(* IEC 61131-3 sources: plc-process-lib/tests/POUs/Suites/FB_DeviceBase_Test, 53 files *)

(* ---- AckAllAcksEveryAlarm.method.decl.st ---- *)
// AckAll() квитирует все тревоги устройства: три активных слота → ActiveAck, wAlmUnack = 0, бит
// DEV_STS_ALARM_UNACK снят, результат Accepted; когда квитировать нечего, AckAll() — FALSE.
// Бит stCmd.xAck делает то же и сбрасывается.
METHOD PRIVATE AckAllAcksEveryAlarm
VAR
    fbTime   : FB_FakeTime;        // подменное время
    fbDev    : FB_TestDevice;      // устройство под тестом
    stCmd    : ST_TestDeviceCmd;   // команды
    stRetain : ST_DeviceRetain;    // энергонезависимые данные
    stCfg    : ST_TestDeviceCfg;   // конфигурация по умолчанию
    itfAlm   : I_Alarm;            // слот через интерфейс
    xRet     : BOOL;               // ответ AckAll
END_VAR

(* ---- AckMaskAcksOnlySelectedSlot.method.decl.st ---- *)
// Маска wAckReq квитирует только выбранный слот (бит 1), маска обнуляется, результат Accepted.
METHOD PRIVATE AckMaskAcksOnlySelectedSlot
VAR
    fbTime   : FB_FakeTime;        // подменное время
    fbDev    : FB_TestDevice;      // устройство под тестом
    stCmd    : ST_TestDeviceCmd;   // команды
    stRetain : ST_DeviceRetain;    // энергонезависимые данные
    stCfg    : ST_TestDeviceCfg;   // конфигурация по умолчанию
    itfAlm   : I_Alarm;            // слот через интерфейс
END_VAR

(* ---- AlarmIdsBaseFromCfgPlusSlot.method.decl.st ---- *)
// Номер тревоги слота = stCfg.udiAlarmIdBase + слот: база 120, слот 5 — 125; номер и значение
// процесса приходят в событии.
METHOD PRIVATE AlarmIdsBaseFromCfgPlusSlot
VAR
    fbTime   : FB_FakeTime;        // подменное время
    fbDev    : FB_TestDevice;      // устройство под тестом
    stCmd    : ST_TestDeviceCmd;   // команды
    stRetain : ST_DeviceRetain;    // энергонезависимые данные
    stCfg    : ST_TestDeviceCfg;   // udiAlarmIdBase = 120
    fbSink   : FB_TestSink;        // приёмник событий
    stEv     : ST_AlarmEvent;      // последнее событие
    itfAlm   : I_Alarm;            // слот через интерфейс
END_VAR

(* ---- AlarmPriorityInvalidCfgErrBit.method.decl.st ---- *)
// Приоритет тревоги вне перечисления (9) не проходит CheckAlarmCfg: бит wCfgErr устройства и
// CheckFunction; исправленный приоритет снимает бит.
METHOD PRIVATE AlarmPriorityInvalidCfgErrBit
VAR
    fbTime   : FB_FakeTime;        // подменное время
    fbDev    : FB_TestDevice;      // устройство под тестом
    stCmd    : ST_TestDeviceCmd;   // команды
    stRetain : ST_DeviceRetain;    // энергонезависимые данные
    stCfg    : ST_TestDeviceCfg;   // слот 3: приоритет 9
    uBad     : U_TestEnumInt;      // число вне перечисления
END_VAR

(* ---- AlarmsInOosAllSlotsOutOfService.method.decl.st ---- *)
// OutOfService устройства — OutOfService у всех используемых слотов (3); в wAlmShelved и wAlmSuppressed их нет
// (ALM-2: вывод из работы виден по eMode), неквитированных нет; после выхода активная тревога снова ActiveUnack.
METHOD PRIVATE AlarmsInOosAllSlotsOutOfService
VAR
    fbTime   : FB_FakeTime;        // подменное время
    fbDev    : FB_TestDevice;      // устройство под тестом
    stCmd    : ST_TestDeviceCmd;   // команды
    stRetain : ST_DeviceRetain;    // энергонезависимые данные
    stCfg    : ST_TestDeviceCfg;   // конфигурация по умолчанию
    itfAlm   : I_Alarm;            // слот через интерфейс
END_VAR

(* ---- AlarmSlotArraysMatchDevAlarmsMax.method.decl.st ---- *)
// Длина массивов слотов базы (afbAlarm, axAlmCond, axAlmSuppress, arAlmValue) равна
// GVL_Const.DEV_ALARMS_MAX: циклы базы идут по константе, тест ловит расхождение, если границу
// запишут числом. Тест читает внутренние переменные базы намеренно — это проверка раскладки.
METHOD PRIVATE AlarmSlotArraysMatchDevAlarmsMax
VAR
    fbDev : FB_TestDevice;   // устройство (вызов не нужен)
    fbAlm : FB_Alarm;        // размер одного слота
END_VAR

(* ---- AlarmSummaryWordsAndPrioUnack.method.decl.st ---- *)
// Сводка тревог: слоты Low, High, Medium активны — ePrioUnack = High; квитирован High — Medium;
// слот Medium вернулся без квитирования — wAlmActive = 2#011, wAlmUnack = 2#101; подавление слота 0
// — бит в wAlmSuppressed (не в wAlmShelved, ALM-2) и снят из wAlmUnack.
METHOD PRIVATE AlarmSummaryWordsAndPrioUnack
VAR
    fbTime   : FB_FakeTime;        // подменное время
    fbDev    : FB_TestDevice;      // устройство под тестом
    stCmd    : ST_TestDeviceCmd;   // команды
    stRetain : ST_DeviceRetain;    // энергонезависимые данные
    stCfg    : ST_TestDeviceCfg;   // приоритеты слотов 0…2
END_VAR

(* ---- AutoToManualBumplessKeepsOutput.method.decl.st ---- *)
// Безударный переход Auto → Manual (хук наследника): работающий механизм продолжает работать.
METHOD PRIVATE AutoToManualBumplessKeepsOutput
VAR
    fbTime   : FB_FakeTime;        // подменное время
    fbDev    : FB_TestDevice;      // устройство под тестом
    stCmd    : ST_TestDeviceCmd;   // команды
    stRetain : ST_DeviceRetain;    // энергонезависимые данные
    stCfg    : ST_TestDeviceCfg;   // конфигурация по умолчанию
END_VAR

(* ---- BeginCycleDtZeroOnFirstCallThenFromTimeSource.method.decl.st ---- *)
// BeginCycle: в первом вызове ltDt = 0; затем — шаг подменного времени (250 мс); при «времени
// назад» — 0 (без переполнения LTIME); дальше снова шаг (100 мс).
METHOD PRIVATE BeginCycleDtZeroOnFirstCallThenFromTimeSource
VAR
    fbTime   : FB_FakeTime;        // подменное время
    fbDev    : FB_TestDevice;      // устройство под тестом
    stCmd    : ST_TestDeviceCmd;   // команды
    stRetain : ST_DeviceRetain;    // энергонезависимые данные
    stCfg    : ST_TestDeviceCfg;   // конфигурация по умолчанию
END_VAR

(* ---- CmdBitsClearedAfterProcessing.method.decl.st ---- *)
// Все импульсные биты и маски stCmd (xSetAuto, xSetManual, xSetOos, xReset, xAck, wAckReq,
// wShelveReq, wUnshelveReq, xStart, xStop) сброшены в том же вызове.
METHOD PRIVATE CmdBitsClearedAfterProcessing
VAR
    fbTime   : FB_FakeTime;        // подменное время
    fbDev    : FB_TestDevice;      // устройство под тестом
    stCmd    : ST_TestDeviceCmd;   // команды
    stRetain : ST_DeviceRetain;    // энергонезависимые данные
    stCfg    : ST_TestDeviceCfg;   // конфигурация по умолчанию
END_VAR

(* ---- CmdResultSeqIncrementsPerCommand.method.decl.st ---- *)
// Каждая обработанная команда пишет eCmdResult и увеличивает uiCmdSeq: в одном вызове режим и пуск
// (в Auto отклонён) — +2, результат последней RejectedMode; Reset и маска shelve без
// принявших слотов — +2, результат RejectedState.
METHOD PRIVATE CmdResultSeqIncrementsPerCommand
VAR
    fbTime   : FB_FakeTime;        // подменное время
    fbDev    : FB_TestDevice;      // устройство под тестом
    stCmd    : ST_TestDeviceCmd;   // команды
    stRetain : ST_DeviceRetain;    // энергонезависимые данные
    stCfg    : ST_TestDeviceCfg;   // слот 0: shelve запрещён
END_VAR

(* ---- ConflictingModeRequestsOosWins.method.decl.st ---- *)
// Одновременные запросы режима (xSetAuto, xSetManual, xSetOos и RequestMode(Auto)) — одна команда:
// побеждает OutOfService; затем xSetAuto вместе с RequestMode(Manual) — побеждает Manual и выводит
// из OutOfService. Импульсы сброшены.
METHOD PRIVATE ConflictingModeRequestsOosWins
VAR
    fbTime   : FB_FakeTime;        // подменное время
    fbDev    : FB_TestDevice;      // устройство под тестом
    stCmd    : ST_TestDeviceCmd;   // команды
    stRetain : ST_DeviceRetain;    // энергонезависимые данные
    stCfg    : ST_TestDeviceCfg;   // конфигурация по умолчанию
    xRet     : BOOL;               // ответ RequestMode
END_VAR

(* ---- DefaultAlarmCfgOfAllTypesPassesCheckAlarmCfg.method.decl.st ---- *)
// Умолчания astAlarm Cfg всех семи устройств и тестового проходят CheckAlarmCfg (инвариант
// генератора для конфигурации тревог); массивы astAlarm из DUT передаются в параметр
// ARRAY[0..GVL_Const.DEV_ALARMS_MAX - 1]. Приоритет 5 и -1 — отказ, 4 (Critical) — норма.
METHOD PRIVATE DefaultAlarmCfgOfAllTypesPassesCheckAlarmCfg
VAR
    fbDev  : FB_TestDevice;         // доступ к CheckAlarmCfg
    stAi   : ST_AnalogInputCfg;     // умолчания AI
    stDi   : ST_DigitalInputCfg;    // умолчания DI
    stMot  : ST_MotorCfg;           // умолчания двигателя
    stVlv  : ST_ValveCfg;           // умолчания арматуры
    stCv   : ST_ControlValveCfg;    // умолчания регулирующего клапана
    stPid  : ST_PidCfg;             // умолчания ПИД
    stTest : ST_TestDeviceCfg;      // умолчания тестового устройства
    stSlot : ST_AlarmCfg;           // копия слота
    uBad   : U_TestEnumInt;         // число вне перечисления
END_VAR

(* ---- DerivedBodyWithoutSuperBaseBodyNotRun.method.decl.st ---- *)
// L1 контракта во время выполнения: у наследника со своим телом без SUPER^ тело базы не
// выполняется само — импульс режима не обработан, FinishCycle не вызван (eDevType = None).
METHOD PRIVATE DerivedBodyWithoutSuperBaseBodyNotRun
VAR
    fbTime   : FB_FakeTime;            // подменное время
    fbNo     : FB_TestDeviceNoSuper;   // наследник без SUPER^
    stCmd    : ST_TestDeviceCmd;       // команды
    stRetain : ST_DeviceRetain;        // энергонезависимые данные
    stCfg    : ST_TestDeviceCfg;       // конфигурация по умолчанию
END_VAR

(* ---- DevTypeSetByHeirReportedInStsCommon.method.decl.st ---- *)
// Тип устройства задаёт наследник в первом вызове, FinishCycle пишет его в stCommon.eDevType;
// до первого вызова — None.
METHOD PRIVATE DevTypeSetByHeirReportedInStsCommon
VAR
    fbTime   : FB_FakeTime;        // подменное время
    fbDev    : FB_TestDevice;      // устройство под тестом
    stCmd    : ST_TestDeviceCmd;   // команды
    stRetain : ST_DeviceRetain;    // энергонезависимые данные
    stCfg    : ST_TestDeviceCfg;   // конфигурация по умолчанию
END_VAR

(* ---- FailureSafeStateResetRules.method.decl.st ---- *)
// Безопасное состояние при отказе: выход снят, Fault, NE 107 Failure, бит wFault, Available =
// FALSE. Reset при действующей причине — RejectedFault; причина ушла — отказ держится до Reset();
// после Reset() выход не включается сам (ручная защёлка снята).
METHOD PRIVATE FailureSafeStateResetRules
VAR
    fbTime   : FB_FakeTime;        // подменное время
    fbDev    : FB_TestDevice;      // устройство под тестом
    stCmd    : ST_TestDeviceCmd;   // команды
    stRetain : ST_DeviceRetain;    // энергонезависимые данные
    stCfg    : ST_TestDeviceCfg;   // конфигурация по умолчанию
    xRet     : BOOL;               // ответ Reset
END_VAR

(* ---- GetAlarmOutOfRangeReturnsNull.method.decl.st ---- *)
// GetAlarm отдаёт слот только в 0..AlarmCount - 1: при трёх слотах — слоты 0…2, номер 3 и 65535 —
// 0; до первого вызова слотов нет.
METHOD PRIVATE GetAlarmOutOfRangeReturnsNull
VAR
    fbTime   : FB_FakeTime;        // подменное время
    fbDev    : FB_TestDevice;      // устройство под тестом
    stCmd    : ST_TestDeviceCmd;   // команды
    stRetain : ST_DeviceRetain;    // энергонезависимые данные
    stCfg    : ST_TestDeviceCfg;   // конфигурация по умолчанию
    itfAlm   : I_Alarm;            // ответ GetAlarm
END_VAR

(* ---- HookViaThisDispatchesToMostDerivedOverride.method.decl.st ---- *)
// Вопрос R2 для двух уровней: у FB_TestDeviceExt хук переопределён ещё раз. THIS^.OnModeChanged из
// метода FB_DeviceBase вызывает реализацию самого производного ФБ; её SUPER^.OnModeChanged
// выполняет часть FB_TestDevice, затем своя часть: след 12 на одну смену режима, 1212 — на две.
METHOD PRIVATE HookViaThisDispatchesToMostDerivedOverride
VAR
    fbTime   : FB_FakeTime;        // подменное время
    fbExt    : FB_TestDeviceExt;   // наследник второго уровня
    stCmd    : ST_TestDeviceCmd;   // команды
    stRetain : ST_DeviceRetain;    // энергонезависимые данные
    stCfg    : ST_TestDeviceCfg;   // конфигурация по умолчанию
END_VAR

(* ---- ImplementsIDeviceInterfaceAccess.method.decl.st ---- *)
// Устройства через I_Device (массив интерфейсов, как у станционной логики): RequestMode, Reset,
// Mode, Status, Fault, Available, AlarmCount, GetAlarm, AckAll работают одинаково для
// FB_TestDevice и его наследника.
METHOD PRIVATE ImplementsIDeviceInterfaceAccess
VAR
    fbTime    : FB_FakeTime;        // подменное время
    fbDev     : FB_TestDevice;      // первое устройство
    fbExt     : FB_TestDeviceExt;   // второе устройство (наследник)
    stCmd     : ST_TestDeviceCmd;   // команды первого
    stRetain  : ST_DeviceRetain;    // retain первого
    stCmd2    : ST_TestDeviceCmd;   // команды второго
    stRetain2 : ST_DeviceRetain;    // retain второго
    stCfg     : ST_TestDeviceCfg;   // общая конфигурация
    aitfDev   : ARRAY[0..1] OF I_Device;   // устройства через интерфейс
    itfDev    : I_Device;           // элемент массива
    itfAlm    : I_Alarm;            // тревога через интерфейс
    uiDev     : UINT;               // номер устройства
    xAllAuto  : BOOL := TRUE;       // все в Auto
    xRet      : BOOL;               // ответы методов
END_VAR

(* ---- ImplementsIDeviceInterfaceAccess.method.impl.st ---- *)
coUnit.TEST('Device_ImplementsIDevice_InterfaceAccess');

aitfDev[0] := fbDev;
aitfDev[1] := fbExt;
FOR uiDev := 0 TO 1 DO
    itfDev := aitfDev[uiDev];
    itfDev.RequestMode(eNewMode := E_DeviceMode.Auto);
END_FOR
fbDev.axCondIn[0] := TRUE;
fbDev(xFaultCause := TRUE, itfTime := fbTime, stCmd := stCmd, stRetain := stRetain, stCfg := stCfg);
fbExt(itfTime := fbTime, stCmd := stCmd2, stRetain := stRetain2, stCfg := stCfg);
FOR uiDev := 0 TO 1 DO
    itfDev := aitfDev[uiDev];
    xAllAuto := xAllAuto AND itfDev.Mode = E_DeviceMode.Auto;
END_FOR
AssertTrue(Condition := xAllAuto, Message := 'RequestMode through the interface');
itfDev := aitfDev[0];
AssertTrue(Condition := itfDev.Fault, Message := 'Fault through the interface');
AssertTrue(Condition := itfDev.Status = E_Ne107Status.Failure, Message := 'Status through the interface');
AssertFalse(Condition := itfDev.Available, Message := 'Available through the interface');
AssertEquals_UINT(Expected := 8, Actual := itfDev.AlarmCount, Message := 'AlarmCount through the interface');
itfAlm := itfDev.GetAlarm(uiIndex := 0);
AssertTrue(Condition := itfAlm.Unacked, Message := 'GetAlarm through the interface');
xRet := itfDev.AckAll();
AssertTrue(Condition := xRet, Message := 'AckAll through the interface');
itfDev.Reset();
fbDev(xFaultCause := FALSE, itfTime := fbTime, stCmd := stCmd, stRetain := stRetain, stCfg := stCfg);
AssertFalse(Condition := itfDev.Fault, Message := 'Reset through the interface');
AssertFalse(Condition := itfAlm.Unacked, Message := 'alarm acknowledged');
itfDev := aitfDev[1];
AssertTrue(Condition := itfDev.Available, Message := 'second device available in Auto');

coUnit.TEST_FINISHED();

(* ---- InputLikeModeMemStartsAutoManualIsCheck.method.decl.st ---- *)
// AI/DI-подобное устройство (без stRetain, режима Local нет): после старта Auto из stModeMem,
// переключатель «Местное» не действует, xSetManual — Manual (подмена) с CheckFunction; stRetain не
// трогается.
METHOD PRIVATE InputLikeModeMemStartsAutoManualIsCheck
VAR
    fbTime   : FB_FakeTime;        // подменное время
    fbIn     : FB_TestDevice;      // устройство под тестом
    stCmd    : ST_TestDeviceCmd;   // команды
    stRetain : ST_DeviceRetain;    // не используется
    stCfg    : ST_TestDeviceCfg;   // конфигурация по умолчанию
END_VAR

(* ---- InvalidCfgAtStartCheckFunctionSafeOutput.method.decl.st ---- *)
// Корректной Cfg ещё не было (rGain = 0): бит wCfgErr, NE 107 CheckFunction, DEV_STS_CFG_ERROR,
// безопасный выход (FALSE и в Auto с запросом), Available = FALSE, пуск — RejectedCfg; режимы
// работают.
METHOD PRIVATE InvalidCfgAtStartCheckFunctionSafeOutput
VAR
    fbTime   : FB_FakeTime;        // подменное время
    fbDev    : FB_TestDevice;      // устройство под тестом
    stCmd    : ST_TestDeviceCmd;   // команды
    stRetain : ST_DeviceRetain;    // энергонезависимые данные
    stCfg    : ST_TestDeviceCfg;   // rGain = 0 — неверно
END_VAR

(* ---- InvalidCfgDuringOperationKeepsLastValidCfg.method.decl.st ---- *)
// Cfg испорчена в работе (rGain = -1): бит wCfgErr и CheckFunction, но логика работает по LKG
// (значение 20 от rGain = 2), механизм не останавливается, Available не меняется; исправленная
// Cfg (rGain = 3) принимается сразу.
METHOD PRIVATE InvalidCfgDuringOperationKeepsLastValidCfg
VAR
    fbTime   : FB_FakeTime;        // подменное время
    fbDev    : FB_TestDevice;      // устройство под тестом
    stCmd    : ST_TestDeviceCmd;   // команды
    stRetain : ST_DeviceRetain;    // энергонезависимые данные
    stCfg    : ST_TestDeviceCfg;   // rGain = 2, затем -1 и 3
END_VAR

(* ---- LocalModeNe107CheckFunction.method.decl.st ---- *)
// Local (переключатель на месте, тип с Local): ПЛК механизмом не управляет — сводный NE 107 CheckFunction («местное
// управление», категория C NE 107, статус PA 0x3C), Available = FALSE; отказ в Local старше — Failure. Возврат в
// дистанционный режим — Good.
METHOD PRIVATE LocalModeNe107CheckFunction
VAR
    fbTime   : FB_FakeTime;        // подменное время
    fbDev    : FB_TestDevice;      // устройство под тестом
    stCmd    : ST_TestDeviceCmd;   // команды
    stRetain : ST_DeviceRetain;    // энергонезависимые данные
    stCfg    : ST_TestDeviceCfg;   // конфигурация
END_VAR

(* ---- LocalOverridesRemoteReturnsToRememberedMode.method.decl.st ---- *)
// Local старше дистанционного режима: в Local выходы сняты, запомненный режим (Auto) сохранён;
// после возврата переключателя устройство продолжает в Auto. Хук — на каждой смене режима.
METHOD PRIVATE LocalOverridesRemoteReturnsToRememberedMode
VAR
    fbTime   : FB_FakeTime;        // подменное время
    fbDev    : FB_TestDevice;      // устройство под тестом
    stCmd    : ST_TestDeviceCmd;   // команды
    stRetain : ST_DeviceRetain;    // энергонезависимые данные
    stCfg    : ST_TestDeviceCfg;   // конфигурация по умолчанию
END_VAR

(* ---- MethodRequestsProcessedOnce.method.decl.st ---- *)
// Запросы методов Reset(), AckAll() и RequestMode() выполняет один ближайший вызов тела, затем они
// снимаются (FinishCycle): uiCmdSeq растёт на 1 за запрос, а не в каждом цикле; тревога, появившаяся
// после выполненного запроса, остаётся неквитированной; режим, сменённый командой после
// RequestMode(), повторный запрос не возвращает. Иначе Reset() станции квитировал бы все будущие
// тревоги и бесконечно повторял бы сброс
METHOD PRIVATE MethodRequestsProcessedOnce
VAR
    fbTime   : FB_FakeTime;        // подменное время
    fbDev    : FB_TestDevice;      // устройство под тестом
    stCmd    : ST_TestDeviceCmd;   // команды
    stRetain : ST_DeviceRetain;    // энергонезависимые данные
    stCfg    : ST_TestDeviceCfg;   // конфигурация по умолчанию
    iStep    : INT;                // шаг цикла
END_VAR

(* ---- MethodRequestsProcessedOnce.method.impl.st ---- *)
coUnit.TEST('Device_MethodRequests_ProcessedOnce');

fbDev(itfTime := fbTime, stCmd := stCmd, stRetain := stRetain, stCfg := stCfg);
fbDev.Reset();
FOR iStep := 1 TO 3 DO
    fbTime.Advance(tStep := T#100MS);
    fbDev(itfTime := fbTime, stCmd := stCmd, stRetain := stRetain, stCfg := stCfg);
END_FOR
AssertEquals_UINT(Expected := 1, Actual := fbDev.stSts.stCommon.uiCmdSeq, Message := 'Reset() executed once');
fbDev.axCondIn[0] := TRUE;
fbDev(itfTime := fbTime, stCmd := stCmd, stRetain := stRetain, stCfg := stCfg);
fbDev(itfTime := fbTime, stCmd := stCmd, stRetain := stRetain, stCfg := stCfg);
AssertEquals_WORD(Expected := 16#0001, Actual := fbDev.stSts.stCommon.wAlmUnack,
                  Message := 'alarm after Reset() stays unacknowledged');
AssertEquals_UINT(Expected := 1, Actual := fbDev.stSts.stCommon.uiCmdSeq, Message := 'no repeated reset');

fbDev.AckAll();
fbDev(itfTime := fbTime, stCmd := stCmd, stRetain := stRetain, stCfg := stCfg);
AssertEquals_WORD(Expected := 0, Actual := fbDev.stSts.stCommon.wAlmUnack, Message := 'AckAll() acknowledged');
fbDev.axCondIn[1] := TRUE;
fbDev(itfTime := fbTime, stCmd := stCmd, stRetain := stRetain, stCfg := stCfg);
fbDev(itfTime := fbTime, stCmd := stCmd, stRetain := stRetain, stCfg := stCfg);
AssertEquals_WORD(Expected := 16#0002, Actual := fbDev.stSts.stCommon.wAlmUnack,
                  Message := 'alarm after AckAll() stays unacknowledged');
AssertEquals_UINT(Expected := 2, Actual := fbDev.stSts.stCommon.uiCmdSeq, Message := 'AckAll() executed once');

fbDev.RequestMode(eNewMode := E_DeviceMode.Auto);
fbDev(itfTime := fbTime, stCmd := stCmd, stRetain := stRetain, stCfg := stCfg);
AssertTrue(Condition := fbDev.Mode = E_DeviceMode.Auto, Message := 'RequestMode(Auto) executed');
stCmd.stCommon.xSetManual := TRUE;
fbDev(itfTime := fbTime, stCmd := stCmd, stRetain := stRetain, stCfg := stCfg);
fbDev(itfTime := fbTime, stCmd := stCmd, stRetain := stRetain, stCfg := stCfg);
AssertTrue(Condition := fbDev.Mode = E_DeviceMode.Manual, Message := 'old RequestMode(Auto) does not come back');
AssertEquals_UINT(Expected := 4, Actual := fbDev.stSts.stCommon.uiCmdSeq, Message := 'four commands in total');

coUnit.TEST_FINISHED();

(* ---- ModeRequestInLocalChangesRememberedMode.method.decl.st ---- *)
// В Local команда xSetAuto принимается и меняет только запомненный режим; после возврата
// переключателя устройство работает в Auto.
METHOD PRIVATE ModeRequestInLocalChangesRememberedMode
VAR
    fbTime   : FB_FakeTime;        // подменное время
    fbDev    : FB_TestDevice;      // устройство под тестом
    stCmd    : ST_TestDeviceCmd;   // команды
    stRetain : ST_DeviceRetain;    // энергонезависимые данные
    stCfg    : ST_TestDeviceCfg;   // конфигурация по умолчанию
END_VAR

(* ---- NoTimeSourceUsesSystemTime.method.decl.st ---- *)
// Без источника (itfTime = 0) база берёт встроенный FB_SystemTime: действующий источник задан,
// время вызова больше 0, шаг между двумя соседними вызовами меньше 1 с.
METHOD PRIVATE NoTimeSourceUsesSystemTime
VAR
    fbDev    : FB_TestDevice;      // устройство под тестом
    stCmd    : ST_TestDeviceCmd;   // команды
    stRetain : ST_DeviceRetain;    // энергонезависимые данные
    stCfg    : ST_TestDeviceCfg;   // конфигурация по умолчанию
END_VAR

(* ---- OnModeChangedHookCalledInDerived.method.decl.st ---- *)
// Вопрос R2 контракта: хук OnModeChanged, вызванный как THIS^.OnModeChanged из метода базы
// (ProcessMode, SwitchRemoteMode), выполняет переопределение наследника с параметрами смены.
METHOD PRIVATE OnModeChangedHookCalledInDerived
VAR
    fbTime   : FB_FakeTime;        // подменное время
    fbDev    : FB_TestDevice;      // устройство под тестом
    stCmd    : ST_TestDeviceCmd;   // команды
    stRetain : ST_DeviceRetain;    // энергонезависимые данные
    stCfg    : ST_TestDeviceCfg;   // конфигурация по умолчанию
END_VAR

(* ---- OosEntryClearsLatchedFaults.method.decl.st ---- *)
// Вход в OutOfService снимает зафиксированные отказы (хук наследника): отказ без Reset держится,
// после xSetOos — Fault = FALSE, статус CheckFunction, wFault = 0; после выхода в Manual — Good.
METHOD PRIVATE OosEntryClearsLatchedFaults
VAR
    fbTime   : FB_FakeTime;        // подменное время
    fbDev    : FB_TestDevice;      // устройство под тестом
    stCmd    : ST_TestDeviceCmd;   // команды
    stRetain : ST_DeviceRetain;    // энергонезависимые данные
    stCfg    : ST_TestDeviceCfg;   // конфигурация по умолчанию
END_VAR

(* ---- OosExitWithLocalSelectedGoesLocal.method.decl.st ---- *)
// OutOfService старше Local: при переключателе «Местное» устройство остаётся OutOfService; выход из
// OutOfService командой xSetManual при включённом «Местном» — в Local.
METHOD PRIVATE OosExitWithLocalSelectedGoesLocal
VAR
    fbTime   : FB_FakeTime;        // подменное время
    fbDev    : FB_TestDevice;      // устройство под тестом
    stCmd    : ST_TestDeviceCmd;   // команды
    stRetain : ST_DeviceRetain;    // энергонезависимые данные
    stCfg    : ST_TestDeviceCfg;   // конфигурация по умолчанию
END_VAR

(* ---- OosRepeatWhileMovingInOosAccepted.method.decl.st ---- *)
// Повтор запроса OutOfService, когда устройство уже выведено из работы, а механизм движется (двигают по месту,
// xMoving): принимается (F-22 (в)) — битом команды и RequestMode: Accepted, uiCmdSeq + 1, режим OutOfService.
METHOD PRIVATE OosRepeatWhileMovingInOosAccepted
VAR
    fbTime   : FB_FakeTime;        // подменное время
    fbDev    : FB_TestDevice;      // устройство под тестом
    stCmd    : ST_TestDeviceCmd;   // команды
    stRetain : ST_DeviceRetain;    // энергонезависимые данные
    stCfg    : ST_TestDeviceCfg;   // конфигурация

    uiSeq    : UINT;               // номер команды после вывода из работы
    xRet     : BOOL;               // ответ RequestMode
END_VAR

(* ---- OutOfServiceRetainedStartsInOos.method.decl.st ---- *)
// stRetain.xOutOfService = TRUE после перезапуска: устройство стартует в OutOfService (хук — в
// первом вызове), все слоты тревог OutOfService; xSetAuto выводит из OutOfService.
METHOD PRIVATE OutOfServiceRetainedStartsInOos
VAR
    fbTime   : FB_FakeTime;        // подменное время
    fbDev    : FB_TestDevice;      // устройство под тестом
    stCmd    : ST_TestDeviceCmd;   // команды
    stRetain : ST_DeviceRetain;    // OutOfService сохранён
    stCfg    : ST_TestDeviceCfg;   // конфигурация по умолчанию
    itfAlm   : I_Alarm;            // слот через интерфейс
END_VAR

(* ---- RequestModeLocalReturnsFalse.method.decl.st ---- *)
// RequestMode(Local) и значение вне перечисления возвращают FALSE: запроса нет, команда не считается.
METHOD PRIVATE RequestModeLocalReturnsFalse
VAR
    fbTime   : FB_FakeTime;        // подменное время
    fbDev    : FB_TestDevice;      // устройство под тестом
    stCmd    : ST_TestDeviceCmd;   // команды
    stRetain : ST_DeviceRetain;    // энергонезависимые данные
    stCfg    : ST_TestDeviceCfg;   // конфигурация по умолчанию
    uBad     : U_TestEnumInt;      // число вне перечисления
    xRet     : BOOL;               // ответы RequestMode
END_VAR

(* ---- RequestModeSameEffectAsCmd.method.decl.st ---- *)
// RequestMode() — запрос, как бит stCmd: режим меняет ближайший вызов тела, результат и uiCmdSeq —
// как у команды; OutOfService при движущемся механизме — RejectedState и через метод, и через бит.
METHOD PRIVATE RequestModeSameEffectAsCmd
VAR
    fbTime   : FB_FakeTime;        // подменное время
    fbDev    : FB_TestDevice;      // устройство под тестом
    stCmd    : ST_TestDeviceCmd;   // команды
    stRetain : ST_DeviceRetain;    // энергонезависимые данные
    stCfg    : ST_TestDeviceCfg;   // конфигурация по умолчанию
    xRet     : BOOL;               // ответ RequestMode
END_VAR

(* ---- ResetCmdAcksAlarmsAndClearsLatch.method.decl.st ---- *)
// stCmd.xReset: сброс зафиксированного отказа (причина ушла) и квитирование всех тревог — одна
// команда (результат Accepted, uiCmdSeq + 1), бит сброшен. Метод Reset() квитирует так же.
METHOD PRIVATE ResetCmdAcksAlarmsAndClearsLatch
VAR
    fbTime   : FB_FakeTime;        // подменное время
    fbDev    : FB_TestDevice;      // устройство под тестом
    stCmd    : ST_TestDeviceCmd;   // команды
    stRetain : ST_DeviceRetain;    // энергонезависимые данные
    stCfg    : ST_TestDeviceCfg;   // конфигурация по умолчанию
    xRet     : BOOL;               // ответ Reset
END_VAR

(* ---- ResolveTimeBeforeBeginCycleNestedDelayDeterministic.method.decl.st ---- *)
// ResolveTime до BeginCycle: вложенный FB_Delay, вызванный раньше BeginCycle, с первого вызова
// получает подменное время — задержка включения 2 с отрабатывает ровно (на 1,9 с выхода нет).
METHOD PRIVATE ResolveTimeBeforeBeginCycleNestedDelayDeterministic
VAR
    fbTime   : FB_FakeTime;        // подменное время
    fbDev    : FB_TestDevice;      // устройство под тестом
    stCmd    : ST_TestDeviceCmd;   // команды
    stRetain : ST_DeviceRetain;    // Auto
    stCfg    : ST_TestDeviceCfg;   // tRunDelay = 2 с
    iStep    : INT;                // шаг цикла
END_VAR

(* ---- ResolveTimeBeforeBeginCycleNestedDelayDeterministic.method.impl.st ---- *)
coUnit.TEST('Device_ResolveTimeBeforeBeginCycle_NestedDelayDeterministic');

stCfg.tRunDelay := T#2S;
stRetain.eRemoteMode := E_DeviceMode.Auto;
fbDev(xAutoRun := FALSE, itfTime := fbTime, stCmd := stCmd, stRetain := stRetain, stCfg := stCfg);   // первый
fbTime.Advance(tStep := T#1S);
fbDev(xAutoRun := TRUE, itfTime := fbTime, stCmd := stCmd, stRetain := stRetain, stCfg := stCfg);    // t1
FOR iStep := 1 TO 19 DO
    fbTime.Advance(tStep := T#100MS);
    fbDev(xAutoRun := TRUE, itfTime := fbTime, stCmd := stCmd, stRetain := stRetain, stCfg := stCfg);
END_FOR
AssertFalse(Condition := fbDev.xOutput, Message := 'no output at t1 + 1.9 s');
fbTime.Advance(tStep := T#100MS);
fbDev(xAutoRun := TRUE, itfTime := fbTime, stCmd := stCmd, stRetain := stRetain, stCfg := stCfg);    // t1 + 2,0 с
AssertTrue(Condition := fbDev.xOutput, Message := 'output exactly at t1 + 2.0 s');

coUnit.TEST_FINISHED();

(* ---- RetainModeInvalidSanitizedToManual.method.decl.st ---- *)
// Значение вне {Auto, Manual} в stRetain.eRemoteMode (7 — мусор, 0 — очищенная память) заменяется
// на Manual и записывается обратно; устройство работает в Manual; это не команда (uiCmdSeq = 0).
METHOD PRIVATE RetainModeInvalidSanitizedToManual
VAR
    fbTime   : FB_FakeTime;        // подменное время
    fbDev    : FB_TestDevice;      // устройство под тестом
    stCmd    : ST_TestDeviceCmd;   // команды
    stRetain : ST_DeviceRetain;    // энергонезависимые данные
    stCfg    : ST_TestDeviceCfg;   // конфигурация по умолчанию
    uBad     : U_TestEnumInt;      // число вне перечисления
END_VAR

(* ---- SetSlotCfg.method.decl.st ---- *)
// Помощник: приоритет и срок shelve слота тревоги в Cfg тестового устройства (через копию элемента)
METHOD PRIVATE SetSlotCfg
VAR_IN_OUT
    stCfgDev : ST_TestDeviceCfg;    // конфигурация устройства
END_VAR
VAR_INPUT
    uiSlot     : UINT;              // номер слота
    ePriority  : E_AlarmPriority;   // приоритет
    tShelveMax : TIME;              // максимальный срок shelve
END_VAR
VAR
    stSlot : ST_AlarmCfg;           // копия слота
END_VAR

(* ---- ShelvedAndSuppressedSeparateMasks.method.decl.st ---- *)
// Отложенная оператором тревога и подавленная логикой — разные биты (ISA-18.2, ALM-2): слот 0 отложен (wShelveReq)
// — бит только в wAlmShelved; слот 1 подавлен (axSuppressIn) — бит только в wAlmSuppressed. Вывод устройства из
// работы — ни shelve, ни подавление: оба слова 0 (OutOfService виден по eMode).
METHOD PRIVATE ShelvedAndSuppressedSeparateMasks
VAR
    fbTime   : FB_FakeTime;        // подменное время
    fbDev    : FB_TestDevice;      // устройство под тестом
    stCmd    : ST_TestDeviceCmd;   // команды
    stRetain : ST_DeviceRetain;    // энергонезависимые данные
    stCfg    : ST_TestDeviceCfg;   // конфигурация
END_VAR

(* ---- ShelveMaskNotAcceptedRejectedState.method.decl.st ---- *)
// Маска shelve, которую не принял ни один слот (у слота tShelveMax = 0; бит неиспользуемого слота),
// даёт результат RejectedState; слот остаётся ActiveUnack.
METHOD PRIVATE ShelveMaskNotAcceptedRejectedState
VAR
    fbTime   : FB_FakeTime;        // подменное время
    fbDev    : FB_TestDevice;      // устройство под тестом
    stCmd    : ST_TestDeviceCmd;   // команды
    stRetain : ST_DeviceRetain;    // энергонезависимые данные
    stCfg    : ST_TestDeviceCfg;   // слот 1: shelve запрещён
    itfAlm   : I_Alarm;            // слот через интерфейс
END_VAR

(* ---- ShelveMaskOnOosEntryRejectedState.method.decl.st ---- *)
// Маска shelve в вызове, в котором устройство уходит в OutOfService (xSetOos и wShelveReq вместе), и
// в OutOfService: shelve не принимается (10.1) — результат маски RejectedState, а не ложный Accepted
// (слот в этот момент ещё не в OutOfService и на запрос ответил бы TRUE); после выхода из
// OutOfService тревога не Shelved
METHOD PRIVATE ShelveMaskOnOosEntryRejectedState
VAR
    fbTime   : FB_FakeTime;        // подменное время
    fbDev    : FB_TestDevice;      // устройство под тестом
    stCmd    : ST_TestDeviceCmd;   // команды
    stRetain : ST_DeviceRetain;    // энергонезависимые данные
    stCfg    : ST_TestDeviceCfg;   // конфигурация по умолчанию (tShelveMax 8 ч)
    itfAlm   : I_Alarm;            // слот 0 через интерфейс
END_VAR

(* ---- ShelveMaskShelvesSlotForMax.method.decl.st ---- *)
// Маска wShelveReq откладывает слот на его tShelveMax (1 ч): Shelved, бит в wAlmShelved, в 50 мин
// ещё отложен, в 60 мин снова ActiveUnack. Маска обнуляется, результат Accepted.
METHOD PRIVATE ShelveMaskShelvesSlotForMax
VAR
    fbTime   : FB_FakeTime;        // подменное время
    fbDev    : FB_TestDevice;      // устройство под тестом
    stCmd    : ST_TestDeviceCmd;   // команды
    stRetain : ST_DeviceRetain;    // энергонезависимые данные
    stCfg    : ST_TestDeviceCfg;   // слот 2: tShelveMax = 1 ч
    itfAlm   : I_Alarm;            // слот через интерфейс
    iStep    : INT;                // шаг цикла
END_VAR

(* ---- ShelveMaskShelvesSlotForMax.method.impl.st ---- *)
coUnit.TEST('Device_ShelveMask_ShelvesSlotForMax');

SetSlotCfg(stCfgDev := stCfg, uiSlot := 2, ePriority := E_AlarmPriority.Medium, tShelveMax := T#1H);
fbDev.axCondIn[2] := TRUE;
fbDev(itfTime := fbTime, stCmd := stCmd, stRetain := stRetain, stCfg := stCfg);
stCmd.stCommon.wShelveReq := 16#0004;
fbDev(itfTime := fbTime, stCmd := stCmd, stRetain := stRetain, stCfg := stCfg);       // t0
itfAlm := fbDev.GetAlarm(uiIndex := 2);
AssertTrue(Condition := itfAlm.State = E_AlarmState.Shelved, Message := 'slot 2 shelved');
AssertEquals_WORD(Expected := 16#0004, Actual := fbDev.stSts.stCommon.wAlmShelved, Message := 'shelved bit');
AssertEquals_WORD(Expected := 0, Actual := fbDev.stSts.stCommon.wAlmUnack, Message := 'no unacknowledged alarm');
AssertEquals_WORD(Expected := 0, Actual := stCmd.stCommon.wShelveReq, Message := 'mask cleared');
AssertTrue(Condition := fbDev.stSts.stCommon.eCmdResult = E_CmdResult.Accepted, Message := 'shelve mask accepted');
FOR iStep := 1 TO 5 DO
    fbTime.Advance(tStep := T#10M);
    fbDev(itfTime := fbTime, stCmd := stCmd, stRetain := stRetain, stCfg := stCfg);
END_FOR
AssertTrue(Condition := itfAlm.State = E_AlarmState.Shelved, Message := 'still shelved at 50 min');
fbTime.Advance(tStep := T#10M);
fbDev(itfTime := fbTime, stCmd := stCmd, stRetain := stRetain, stCfg := stCfg);       // t0 + 1 ч
AssertTrue(Condition := itfAlm.State = E_AlarmState.ActiveUnack, Message := 'reannunciated after tShelveMax');
AssertEquals_WORD(Expected := 0, Actual := fbDev.stSts.stCommon.wAlmShelved, Message := 'shelved bit cleared');

coUnit.TEST_FINISHED();

(* ---- StopInAutoSwitchesToManual.method.decl.st ---- *)
// «Стоп» оператора в Auto: SwitchRemoteMode переводит в Manual сразу (хук Auto → Manual), режим
// записан в retain, механизм остановлен, результат Accepted.
METHOD PRIVATE StopInAutoSwitchesToManual
VAR
    fbTime   : FB_FakeTime;        // подменное время
    fbDev    : FB_TestDevice;      // устройство под тестом
    stCmd    : ST_TestDeviceCmd;   // команды
    stRetain : ST_DeviceRetain;    // энергонезависимые данные
    stCfg    : ST_TestDeviceCfg;   // конфигурация по умолчанию
END_VAR

(* ---- StsHeaderAllFieldsFilled.method.decl.st ---- *)
// FinishCycle заполняет все 14 полей stCommon: слово состояния (биты устройства и общие),
// wFault, wWarning, wCfgErr, режим, NE 107, результат и номер команды, маски тревог, наивысший
// приоритет неквитированных, тип устройства, резерв.
METHOD PRIVATE StsHeaderAllFieldsFilled
VAR
    fbTime   : FB_FakeTime;        // подменное время
    fbDev    : FB_TestDevice;      // устройство под тестом
    stCmd    : ST_TestDeviceCmd;   // команды
    stRetain : ST_DeviceRetain;    // энергонезависимые данные
    stCfg    : ST_TestDeviceCfg;   // слот 0: High
    stHdr    : ST_DeviceSts;       // копия заголовка
END_VAR

(* ---- SummaryStatusMaxOfDeviceModeAndCfg.method.decl.st ---- *)
// Сводный NE 107 = MAX(устройство, режим, Cfg): S и M от устройства (бит предупреждения), M при
// испорченной Cfg — C, F в OutOfService — F (Fault, бит отказа), Good в OutOfService — C;
// AI/DI-подобное устройство: Manual (подмена) — C.
METHOD PRIVATE SummaryStatusMaxOfDeviceModeAndCfg
VAR
    fbTime     : FB_FakeTime;        // подменное время
    fbDev      : FB_TestDevice;      // устройство под тестом
    stCmd      : ST_TestDeviceCmd;   // команды
    stRetain   : ST_DeviceRetain;    // энергонезависимые данные
    stCfg      : ST_TestDeviceCfg;   // конфигурация
    fbIn       : FB_TestDevice;      // AI/DI-подобное устройство
    stCmdIn    : ST_TestDeviceCmd;   // его команды
    stRetainIn : ST_DeviceRetain;    // его retain (не используется)
END_VAR

(* ---- SuperBodyCallRunsBaseBodyOnSameStructs.method.decl.st ---- *)
// Вопрос R3 контракта: SUPER^(stCmd := stCmd, stRetain := stRetain, stCfg := stCfg) в теле
// наследника выполняет тело базы один раз за вызов над теми же структурами, что переданы в вызов
// наследника: импульс сброшен и режим записан в структурах вызывающего, Cfg вызывающего прочитана,
// запись наследника в stCmd после SUPER^ видна; точка расширения до SUPER^ действует; вызов с
// другими структурами работает с ними.
METHOD PRIVATE SuperBodyCallRunsBaseBodyOnSameStructs
VAR
    fbTime    : FB_FakeTime;        // подменное время
    fbExt     : FB_TestDeviceExt;   // наследник с SUPER^
    stCmd     : ST_TestDeviceCmd;   // команды (первый набор)
    stRetain  : ST_DeviceRetain;    // энергонезависимые данные (первый набор)
    stCmd2    : ST_TestDeviceCmd;   // команды (второй набор)
    stRetain2 : ST_DeviceRetain;    // энергонезависимые данные (второй набор)
    stCfg     : ST_TestDeviceCfg;   // rGain = 3
END_VAR

(* ---- SwitchRemoteModeInLocalOnlyRemembers.method.decl.st ---- *)
// SwitchRemoteMode в Local меняет только запомненный режим, без смены режима и хука; после возврата
// переключателя — Manual.
METHOD PRIVATE SwitchRemoteModeInLocalOnlyRemembers
VAR
    fbTime   : FB_FakeTime;        // подменное время
    fbDev    : FB_TestDevice;      // устройство под тестом
    stCmd    : ST_TestDeviceCmd;   // команды
    stRetain : ST_DeviceRetain;    // энергонезависимые данные
    stCfg    : ST_TestDeviceCfg;   // конфигурация по умолчанию
    uiHooks  : UINT;               // вызовов хука до SwitchRemoteMode
END_VAR

(* ---- ZeroAlarmCountNoSlotsRun.method.decl.st ---- *)
// Устройство без тревог (uiAlarmCount = 0): все условия и маски взведены — ни один слот не
// вызывается, сводка пустая, GetAlarm(0) = 0; маска квитирования — Accepted, маска shelve —
// RejectedState. Проверка цикла FOR 1 TO MIN(...) без беззнакового «0 - 1».
METHOD PRIVATE ZeroAlarmCountNoSlotsRun
VAR
    fbTime   : FB_FakeTime;        // подменное время
    fbDev    : FB_TestDevice;      // устройство под тестом
    stCmd    : ST_TestDeviceCmd;   // команды
    stRetain : ST_DeviceRetain;    // энергонезависимые данные
    stCfg    : ST_TestDeviceCfg;   // конфигурация по умолчанию
    itfAlm   : I_Alarm;            // ответ GetAlarm
    uiSlot   : UINT;               // номер слота
END_VAR

(* ---- ZeroAlarmCountNoSlotsRun.method.impl.st ---- *)
coUnit.TEST('Device_ZeroAlarmCount_NoSlotsRun');

FOR uiSlot := 0 TO 7 DO
    fbDev.axCondIn[uiSlot] := TRUE;
END_FOR
stCmd.stCommon.wAckReq := 16#FFFF;
fbDev(uiAlarmSlots := 0, itfTime := fbTime, stCmd := stCmd, stRetain := stRetain, stCfg := stCfg);
AssertEquals_UINT(Expected := 0, Actual := fbDev.AlarmCount, Message := 'no alarm slots');
AssertEquals_WORD(Expected := 0, Actual := fbDev.stSts.stCommon.wAlmActive, Message := 'no active alarms');
AssertEquals_WORD(Expected := 0, Actual := fbDev.stSts.stCommon.wAlmUnack, Message := 'no unacknowledged alarms');
AssertTrue(Condition := fbDev.stSts.stCommon.eCmdResult = E_CmdResult.Accepted, Message := 'ack mask accepted');
itfAlm := fbDev.GetAlarm(uiIndex := 0);
AssertTrue(Condition := itfAlm = 0, Message := 'GetAlarm(0) = 0');
stCmd.stCommon.wShelveReq := 16#FFFF;
fbDev(itfTime := fbTime, stCmd := stCmd, stRetain := stRetain, stCfg := stCfg);
AssertTrue(Condition := fbDev.stSts.stCommon.eCmdResult = E_CmdResult.RejectedState,
           Message := 'shelve mask: no slot accepted');

coUnit.TEST_FINISHED();
